(*
SPDX-FileCopyrightText: © 2026 Oleksandr Tiutyk <trofimich@gmail.com>
SPDX-License-Identifier: MIT
License: https://opensource.org/license/mit
*)

(*!
<summary>Exercises the production Task lifecycle with delayed, interruptible stopping.</summary>
<description>
The scenario owns and injects a TaskStoppingResource through SetResource before Start. The binding is borrowed
and stable across runs. Inputs configure faults; ThrowOnEveryStopping may be cleared while RUNNING to resume
cleanup. Observations are cumulative until ClearObservations, except cleanup progress, which OnReset clears.
No physical I/O is performed.
</description>
*)

FUNCTION_BLOCK TaskStoppingProbe EXTENDS TOF_Tasks.Task
VAR_INPUT
	//! <summary>Ordinary OnRunning result when no exception is injected.</summary>
	ProcessingResult : TOF_Tasks.TASK_PROCESSING_STATE := TOF_Tasks.TASK_PROCESSING_STATE.DONE;
	//! <summary>Throw from start preparation before RUNNING is entered.</summary>
	ThrowOnBeforeStart : BOOL;
	//! <summary>Throw when ordinary processing is called.</summary>
	ThrowOnRunning : BOOL;
	//! <summary>Throw once in stopping before advancing cleanup.</summary>
	ThrowOnFirstStopping : BOOL;
	//! <summary>Throw on every stopping call while enabled, before advancing cleanup.</summary>
	ThrowOnEveryStopping : BOOL;
	//! <summary>Throw from reset before descendant state is cleared.</summary>
	ThrowOnReset : BOOL;
	//! <summary>Injected exceptions throw again from GetMessage.</summary>
	ThrowOnGetMessage : BOOL;
	//! <summary>Throw a StandardException whose GetMessage result is empty.</summary>
	ThrowWithEmptyMessage : BOOL;
	//! <summary>Exercise the permitted Reset notification after termination.</summary>
	ResetOnAfterStop : BOOL;
END_VAR
VAR_OUTPUT
	//! <summary>Total ordinary processing calls across runs.</summary>
	RunningCalls : UINT;
	//! <summary>Total stopping-hook calls across runs, including interrupted calls.</summary>
	StoppingCalls : UINT;
	//! <summary>Successful stopping steps since the last Reset.</summary>
	CompletedCleanupSteps : UINT;
	//! <summary>Total notifications after STOPPED has been recorded.</summary>
	AfterStopCalls : UINT;
	//! <summary>Total accepted cancellation notifications.</summary>
	CancelNotifications : UINT;
END_VAR
VAR CONSTANT
	//! <summary>Successful cleanup steps required before release is safe.</summary>
	_CleanupSteps : UINT := 2;
END_VAR
VAR_STAT
	//! <summary>Class name shared by all instances of this function block.</summary>
	_ClassName : STRING := __POUNAME();
END_VAR
VAR
	_Resource : REFERENCE TO TaskStoppingResource;
	_StoppingExceptionRaised : BOOL;
END_VAR

{attribute 'monitoring' := 'call'}
PROPERTY ClassName : REFERENCE TO STRING
GET
ClassName REF= _ClassName;
END_GET
END_PROPERTY

(*!
<summary>Starts a fresh set of observation counts.</summary>
<description>
Call while the fixture is READY. Leaves configuration, cleanup progress and the borrowed resource binding intact.
</description>
*)
METHOD INTERNAL ClearObservations
RunningCalls := 0;
StoppingCalls := 0;
AfterStopCalls := 0;
CancelNotifications := 0;
END_METHOD

(*!
<summary>Borrows the test namespace.</summary>
*)
{attribute 'monitoring' := 'call'}
PROPERTY NamespaceName : REFERENCE TO STRING
GET
NamespaceName REF= CurrentNamespace.Name;
END_GET
END_PROPERTY

(*!
<summary>Counts finalization and optionally resets the stopped task.</summary>
<description>
Reset is invoked only after STOPPED and final diagnostics have been published.
</description>
*)
METHOD PROTECTED OnAfterStop
AfterStopCalls := AfterStopCalls + 1;

IF ResetOnAfterStop THEN
	Reset();
END_IF
END_METHOD

(*!
<summary>Optionally refuses start through an injected exception.</summary>
*)
METHOD PROTECTED OnBeforeStart
IF ThrowOnBeforeStart THEN
	raiseConfiguredFailure(message := "Start failure");
END_IF
END_METHOD

(*!
<summary>Counts accepted external cancellation notifications.</summary>
*)
METHOD PROTECTED OnCancelRequest
CancelNotifications := CancelNotifications + 1;
END_METHOD

(*!
<summary>Clears per-run cleanup progress without resetting observations or the dependency.</summary>
<description>
An injected exception refuses Reset before changing descendant state.
</description>
*)
METHOD PROTECTED OnReset
IF ThrowOnReset THEN
	raiseConfiguredFailure(message := "Reset failure");
END_IF

CompletedCleanupSteps := 0;
_StoppingExceptionRaised := FALSE;
END_METHOD

(*!
<summary>Returns the configured work result or injects a processing exception.</summary>
<description>
One call records one unit of work; no resource operations are driven here.
</description>
<param name="processingState">Configured result on normal return.</param>
<param name="stopReasonMessage">Receives diagnostic text for ERROR or ABORTED.</param>
*)
METHOD PROTECTED OnRunning
VAR_OUTPUT
	processingState : TOF_Tasks.TASK_PROCESSING_STATE;
END_VAR
VAR_IN_OUT
	stopReasonMessage : TOF_Core.ERROR_MESSAGE;
END_VAR
RunningCalls := RunningCalls + 1;

IF ThrowOnRunning THEN
	raiseConfiguredFailure(message := "Work failure");
END_IF

processingState := ProcessingResult;

IF processingState = TOF_Tasks.TASK_PROCESSING_STATE.ERROR
	OR_ELSE processingState = TOF_Tasks.TASK_PROCESSING_STATE.ABORTED
THEN
	stopReasonMessage := "Work result";
END_IF
END_METHOD

(*!
<summary>Finishes late acquisition and two cleanup steps before allowing release.</summary>
<description>
The configured exception can interrupt one or every call before progress. A later call resumes without
rerunning ordinary work once repeated injection is disabled.
</description>
<param name="readyToRelease">TRUE only after pending acquisition and cleanup have completed.</param>
*)
METHOD PROTECTED OnStopping
VAR_OUTPUT
	readyToRelease : BOOL;
END_VAR
StoppingCalls := StoppingCalls + 1;

IF ThrowOnFirstStopping AND_THEN NOT _StoppingExceptionRaised THEN
	_StoppingExceptionRaised := TRUE;
	raiseConfiguredFailure(message := "Stopping failure");
END_IF

IF ThrowOnEveryStopping THEN
	raiseConfiguredFailure(message := "Stopping failure");
END_IF

IF __ISVALIDREF(_Resource) AND_THEN NOT _Resource.FinishPendingAcquire() THEN
	RETURN;
END_IF

CompletedCleanupSteps := CompletedCleanupSteps + 1;
readyToRelease := CompletedCleanupSteps >= _CleanupSteps;
END_METHOD

(*!
<summary>Raises the configured synthetic exception.</summary>
<description>
Used only by test operations, never by FB lifecycle methods. A throwing or empty formatter exercises
diagnostic fallback.
</description>
<param name="message">Text copied into the injected exception.</param>
*)
METHOD PRIVATE raiseConfiguredFailure
VAR_INPUT
	message : WSTRING(255);
END_VAR
VAR
	failure : TOF_Core.StandardException;
	formattingFailure : ThrowingGetMessageException;
	emptyMessage : TOF_Core.ERROR_MESSAGE;
END_VAR
IF ThrowOnGetMessage THEN
	formattingFailure.Throw(
		sourceNamespaceName := NamespaceName,
		sourceClassName := ClassName,
		sourcePOUName := __POUNAME(),
		sourcePosition := __POSITION(),
		message := message
	);
ELSIF ThrowWithEmptyMessage THEN
	emptyMessage := TOF_Core.WideStrings.Empty;
	failure.Throw(
		sourceNamespaceName := NamespaceName,
		sourceClassName := ClassName,
		sourcePOUName := __POUNAME(),
		sourcePosition := __POSITION(),
		message := emptyMessage
	);
ELSE
	failure.Throw(
		sourceNamespaceName := NamespaceName,
		sourceClassName := ClassName,
		sourcePOUName := __POUNAME(),
		sourcePosition := __POSITION(),
		message := message
	);
END_IF
END_METHOD

(*!
<summary>Returns the explicitly injected borrowed resource manager.</summary>
<description>
Zero before binding; getter has no side effects and does not throw.
</description>
*)
{attribute 'monitoring' := 'call'}
PROPERTY ResourceManager : TOF_Core.IResourceManager
GET
IF __ISVALIDREF(_Resource) THEN
	ResourceManager := _Resource;
END_IF
END_GET
END_PROPERTY

(*!
<summary>Reports the concrete fixture size.</summary>
*)
{attribute 'monitoring' := 'call'}
PROPERTY SelfSize : ULINT
GET
SelfSize := XSIZEOF(THIS^);
END_GET
END_PROPERTY

(*!
<summary>Binds the manager owned by the scenario.</summary>
<description>
Call before Start and keep the referenced manager alive and unchanged throughout every run. Reset preserves
the binding.
</description>
<param name="resource">Live synthetic manager owned directly by the scenario.</param>
*)
METHOD INTERNAL SetResource
VAR_IN_OUT
	resource : TaskStoppingResource;
END_VAR
_Resource REF= resource;
END_METHOD

END_FUNCTION_BLOCK

(* stored: Version 1.1.0.1, ProductVersion 3.1.4026.21
   POU TaskStoppingProbe: Id {4e5922b3-4fc0-4824-ba95-5762e94466c9}, SpecialFunc None
   Folder Overriden methods: Id {58e70026-eeaf-4d30-88ef-971ac03e0916}
   Folder Service methods: Id {00187476-6411-4e2f-8536-12a37d7ec040}
   Property ClassName: Id {2c3e4e2a-7f6e-442a-ae42-79e6fbb82217}
   Get Get: Id {f5a6f232-e55c-4d3c-9948-0e2873d9665f}
   Method ClearObservations: Id {5bc1d808-cf80-4464-bb40-9a61d96f4bd6}
   Property NamespaceName: Id {d32ccf65-dbcc-455d-910f-9bcab73d5d17}
   Get Get: Id {2517d35b-1677-487a-a4e0-d8c211d58e02}
   Method OnAfterStop: Id {3beb56c7-ded4-4afc-9026-79e0def1e6ee}
   Method OnBeforeStart: Id {42f11eb6-f2bb-4dba-bbbe-d0bc202bfe7e}
   Method OnCancelRequest: Id {c87816ab-1306-44ac-8f29-45823512d900}
   Method OnReset: Id {ded75715-8c86-4040-bced-7496d56004f2}
   Method OnRunning: Id {9a2dcb9f-4f91-45be-8232-0869e1f5baf0}
   Method OnStopping: Id {a9ea76b2-4078-49f6-a27e-6ecea9963c7d}
   Method raiseConfiguredFailure: Id {76c8b4a3-202c-4375-897d-fe0c747ff965}
   Property ResourceManager: Id {69c0e752-f6a8-45f7-bb1f-89c64b06b3eb}
   Get Get: Id {366116c5-2b57-41a8-8abb-105c25397dc3}
   Property SelfSize: Id {4526353b-c0db-4703-b1dc-9d9b39ec7e72}
   Get Get: Id {145f273b-c5fb-428b-b735-54de013ffc5b}
   Method SetResource: Id {6d4e1126-9421-46d6-b682-23a7a6067960} *)
